// TwinCAT 3 PLC project FixturePlc
// ProgramVersion: 3.1.4026.22
// libraries:
//   Tc2_Standard, * (Beckhoff Automation GmbH)
//   Tc2_System, * (Beckhoff Automation GmbH)
// project tree:
//   DUTs/ E_FixtureMode.TcDUT, ST_FixtureRecord.TcDUT, ST_PersistentInner.TcDUT, ST_PersistentRecipe.TcDUT, T_FixtureName.TcDUT
//   GVLs/ GVL_Fixture.TcGVL, GVL_IBN_Probe.TcGVL, GVL_InstanceSettings.TcGVL, GVL_Persistent.TcGVL
//   / PlcTask.TcTTO
//   POUs/ FB_FolderMembers.TcPOU, FB_PersistentCell.TcPOU, FB_StepChain.TcPOU, I_FixtureDevice.TcIO, MAIN.TcPOU, PRG_IntegrationScratch.TcPOU
// real-time tasks:
//   TASK PlcTask: cycle T#10ms, priority 20, ADS port 350
// motion (NC):
//   TASK NC-Task 1 SAF: cycle T#2ms, priority 4, ADS port 501
//   TASK NC-Task 1 SVB: cycle T#10ms, priority 8, ADS port 511
// I/O:
//   DEVICE Device 1 (EtherCAT) (disabled), AmsNetId 199.4.42.250.2.1
//     Term 1 (EK1100) [EK1100 EtherCAT-Koppler (2A E-Bus)]
//       Term 2 (EL1008) [EL1008 8K. Dig. Eingang 24V, 3ms]
//       Term 3 (EL3174) [EL3174 4K. Ana. Eingang  +/-10V Diff., +/-20mA SingleEnded, 16 Bit]
// variable links:
//   FixturePlc/FixturePlc Instance <-> Device 1 (EtherCAT)/Term 1 (EK1100)/Term 2 (EL1008)
//     PlcTask Inputs/GVL_Fixture.bInputSignal <-> Channel 1/Input

CONFIGURATION FixturePlc
    RESOURCE PLC ON TwinCAT3
        TASK PlcTask(INTERVAL := T#10ms, PRIORITY := 20);
        PROGRAM MAIN WITH PlcTask : MAIN;
    END_RESOURCE
END_CONFIGURATION

// ---- DUTs/E_FixtureMode.TcDUT
{attribute 'qualified_only'}
{attribute 'strict'}
TYPE E_FixtureMode :
(
	Idle := 0,
	Running := 1,
	Done := 2
) INT;
END_TYPE

// ---- DUTs/ST_FixtureRecord.TcDUT
TYPE ST_FixtureRecord :
STRUCT
	nId : UDINT;
	fValue : LREAL;
	sLabel : STRING(40);
	eMode : E_FixtureMode;
END_STRUCT
END_TYPE

// ---- DUTs/ST_PersistentInner.TcDUT
TYPE ST_PersistentInner :
STRUCT
	nCount : INT;
	fOffset : LREAL;
END_STRUCT
END_TYPE

// ---- DUTs/ST_PersistentRecipe.TcDUT
TYPE ST_PersistentRecipe :
STRUCT
	stInner : ST_PersistentInner;
	eMode : E_FixtureMode;
	sName : STRING(20);
	wsName : WSTRING(20);
	tDelay : TIME := T#1S500MS;
	dtStamp : DT;
	aPos : ARRAY[1..5] OF LREAL;
END_STRUCT
END_TYPE

// ---- DUTs/T_FixtureName.TcDUT
TYPE T_FixtureName : STRING(40); END_TYPE

// ---- GVLs/GVL_Fixture.TcGVL
{attribute 'qualified_only'}
VAR_GLOBAL
	bEnable : BOOL;
	bInputSignal AT %I* : BOOL;
	nCount : UINT := 2;
	nCycleCount : UDINT;
	fValue : LREAL := 1.5;
	sText : STRING := 'fixture';
	aNames : ARRAY[0..3] OF STRING(20) := ['alpha', 'beta', 'gamma', 'delta'];
END_VAR

// ---- GVLs/GVL_IBN_Probe.TcGVL
{attribute 'qualified_only'}
VAR_GLOBAL
	bEnable : BOOL; // heartbeat: TRUE while armed, FALSE on disarm/abort/release_all
	bStepReq : BOOL; // the single command bit, written only by a human-confirmed proposal
	bAbort : BOOL; // panic/home: TRUE on disarm/abort/release_all
	bChainRunning : BOOL; // status read by twincat_list_active_chains
	nActiveChain : INT;
	nCurrentStep : INT;
	bFault : BOOL;
END_VAR

// ---- GVLs/GVL_InstanceSettings.TcGVL
{attribute 'qualified_only'}
VAR_GLOBAL
	{attribute 'TcInitSymbol'}
	nInitParam : DINT := 10;
	{attribute 'TcInitSymbol'}
	fInitGain : LREAL := 1.5;
END_VAR
VAR_GLOBAL RETAIN
	nRetainCounter : UDINT;
END_VAR

// ---- GVLs/GVL_Persistent.TcGVL
{attribute 'qualified_only'}
VAR_GLOBAL PERSISTENT
	stRecipe : ST_PersistentRecipe;
	arCal : ARRAY[1..3] OF ST_PersistentInner;
END_VAR
VAR_GLOBAL
	fbCell : FB_PersistentCell;
	aCells : ARRAY[1..2] OF FB_PersistentCell;
END_VAR

// ---- POUs/I_FixtureDevice.TcIO
INTERFACE I_FixtureDevice

METHOD Reset : BOOL
VAR_INPUT
END_VAR
END_METHOD

END_INTERFACE

// ---- POUs/MAIN.TcPOU
PROGRAM MAIN
VAR
	fbStepChain : FB_StepChain;
	stRecord : ST_FixtureRecord;
	eMode : E_FixtureMode;
	sName : T_FixtureName := 'fixture';
	bInput : BOOL;
	sFirstName : STRING(20);
	bIbnProbeIdle : BOOL;
	fInstanceProbe : LREAL;
	stRecipeProbe : ST_PersistentRecipe;
	arCalProbe : ARRAY[1..3] OF ST_PersistentInner;
END_VAR

fbStepChain(bStart := GVL_Fixture.bEnable);
GVL_Fixture.nCycleCount := GVL_Fixture.nCycleCount + 1;
GVL_Fixture.fValue := GVL_Fixture.fValue + 0.001;
bInput := GVL_Fixture.bInputSignal;
sFirstName := GVL_Fixture.aNames[0];
stRecord.nId := GVL_Fixture.nCount;
stRecord.fValue := GVL_Fixture.fValue;
stRecord.sLabel := GVL_Fixture.sText;
stRecord.eMode := eMode;

// IbnLive probe: only read here, so every GVL_IBN_Probe symbol stays in the ADS symbol table.
bIbnProbeIdle := NOT (GVL_IBN_Probe.bEnable OR GVL_IBN_Probe.bStepReq OR GVL_IBN_Probe.bAbort
	OR GVL_IBN_Probe.bChainRunning OR GVL_IBN_Probe.bFault)
	AND GVL_IBN_Probe.nActiveChain = 0 AND GVL_IBN_Probe.nCurrentStep = 0;

// plc-instance-settings: only read here, so the init symbols and the retain variable stay in the image.
fInstanceProbe := GVL_InstanceSettings.fInitGain * DINT_TO_LREAL(GVL_InstanceSettings.nInitParam)
	+ UDINT_TO_LREAL(GVL_InstanceSettings.nRetainCounter);

// persistent-snapshot: the remanent symbols are read here so they stay in the image and the ADS symbol table.
GVL_Persistent.fbCell();
GVL_Persistent.aCells[1]();
GVL_Persistent.aCells[2]();
stRecipeProbe := GVL_Persistent.stRecipe;
arCalProbe := GVL_Persistent.arCal;

PRG_IntegrationScratch(); // [INTEGRATION-TEST-HOOK] do not remove manually

END_PROGRAM

// ---- POUs/FB_StepChain.TcPOU
FUNCTION_BLOCK FB_StepChain
VAR_INPUT
	bStart : BOOL;
END_VAR
VAR
	Step : INT;
	tonWait : TON;
	nRuns : UDINT;
END_VAR

CASE Step OF
	0: // idle
		IF bStart THEN
			Step := 10;
		END_IF

	10: // wait a moment
		tonWait(IN := TRUE, PT := T#100MS);
		IF tonWait.Q THEN
			tonWait(IN := FALSE);
			Step := 1010;
		END_IF

	// 20: commented-out step, must never match

	1010: // work
		nRuns := nRuns + 1;
		Step := 1020;

	1020, 1030: // finish
		Step := 0;

ELSE
	Step := 0;
END_CASE

END_FUNCTION_BLOCK

// ---- POUs/PRG_IntegrationScratch.TcPOU
PROGRAM PRG_IntegrationScratch
VAR
END_VAR

; // integration-test scratch POU. Body is freely overwritten and restored by the live test suite. Never put real logic here.

END_PROGRAM

// ---- POUs/FB_PersistentCell.TcPOU
FUNCTION_BLOCK FB_PersistentCell
VAR PERSISTENT
	nPersistentCount : DINT;
END_VAR
VAR RETAIN
	nRetainCount : DINT;
END_VAR
VAR
	nTransient : DINT;
END_VAR

nTransient := nPersistentCount + nRetainCount;

END_FUNCTION_BLOCK

// ---- POUs/FB_FolderMembers.TcPOU
FUNCTION_BLOCK FB_FolderMembers
VAR_INPUT
END_VAR
VAR_OUTPUT
END_VAR
VAR
END_VAR

PROPERTY PUBLIC Enabled : BOOL
GET // PUBLIC
END_GET
SET // PUBLIC
END_SET
END_PROPERTY

METHOD Reset : BOOL
END_METHOD

END_FUNCTION_BLOCK
